// TIA Portal V21 export
// export: Created 2026-10-23T20:43:16.2360317Z, ExportSetting WithDefaults, DisplayName Totally Integrated Automation Portal, DisplayVersion V21 Update 1, DisplayName SINAMICS Startdrive Advanced, DisplayVersion V21 HF2, DisplayName SINAMICS Startdrive G110M, G120, G120C, G120D, G120P, G115D, DisplayVersion V21 HF2, DisplayName SINAMICS Startdrive G130, G150, S120, S150, G200, G220, S200, S210, S220, Innomotics MVD, DisplayVersion V21 HF2, DisplayName STEP 7 Professional, DisplayVersion V21 Update 1, DisplayName STEP 7 Safety, DisplayVersion V21, DisplayName Tech WebApplication, DisplayVersion V21, DisplayName WinCC Basic/Comfort/Advanced, DisplayVersion V21 Update 1, DisplayName WinCC Unified, DisplayVersion V21 Update 1
FUNCTION "FC_AnaOutputPath" : Void   // FC11, SCL
TITLE = Analyzer: output not written on every path
{ S7_Optimized_Access := 'TRUE' }
VERSION : 0.1
// Rule C26d: Result is not written when Select is FALSE
// stored: AutoNumber true, IsIECCheckEnabled false, SetENOAutomatically false, UDAEnableTagReadback false
   VAR_INPUT
      Select : Bool;   // Select the value
      Value : Int;   // Value
   END_VAR
   VAR_OUTPUT
      Result : Int;   // Result
   END_VAR
BEGIN

       IF #Select THEN
           #Result := #Value;
       END_IF;
END_FUNCTION
